(* PLC project TBEN_L5_PLC11.project, CODESYS CODESYS V3.5 SP21 Patch 1 *)
(* stored: creationDateTime 2026-11-07T15:34:51.4878878, modificationDateTime 2026-11-07T15:09:07.4034196 *)

{attribute 'qualified_only'}
// Loại event IO-Link (= bit 5..4 của EventQualifier)
TYPE E_IolEvtType :
(
    NOTIFICATION := 1,
    WARNING      := 2,
    ERROR        := 3
) INT;
END_TYPE
